(* IEC 61131-3 sources: Test-Git_ESME26/TestProgettoESME_26.fbsproj/AxisModuleLib Migration/DiagSource, 7 files *)

(* ---- AXM_FC_EtCamTypeToString.fn.st ---- *)
FUNCTION INTERNAL AXM_FC_EtCamTypeToString : STRING[80]
VAR_INPUT
	i_etCamType	: CMT.ET_CamType;
END_VAR
VAR
END_VAR

CASE i_etCamType OF
	CMT.ET_CamType.Straight:
		AXM_FC_EtCamTypeToString := 'Straight';

	CMT.ET_CamType.Poly5Com:
		AXM_FC_EtCamTypeToString := 'Poly5Com';

	CMT.ET_CamType.SimplSin:
		AXM_FC_EtCamTypeToString := 'SimplSin';

	CMT.ET_CamType.IncliSin:
		AXM_FC_EtCamTypeToString := 'IncliSin';

	CMT.ET_CamType.ModiSin:
		AXM_FC_EtCamTypeToString := 'ModiSin';

	CMT.ET_CamType.ModAccTr:
		AXM_FC_EtCamTypeToString := 'ModAccTr';

	CMT.ET_CamType.Poly5:
		AXM_FC_EtCamTypeToString := 'Poly5';

	CMT.ET_CamType.Parable2:
		AXM_FC_EtCamTypeToString := 'Parable2';

	CMT.ET_CamType.UserCam:
		AXM_FC_EtCamTypeToString := 'UserCam';

	CMT.ET_CamType.ModiSinCom:
		AXM_FC_EtCamTypeToString := 'ModiSinCom';

	CMT.ET_CamType.ModAccTrCom:
		AXM_FC_EtCamTypeToString := 'ModAccTrCom';

	CMT.ET_CamType.HarmoComb:
		AXM_FC_EtCamTypeToString := 'HarmoComb';

	CMT.ET_CamType.SinStraightComb:
		AXM_FC_EtCamTypeToString := 'SinStraightComb';

ELSE
	AXM_FC_EtCamTypeToString := Standard.CONCAT('Unknown CamType ', INT_TO_STRING(i_etCamType));
END_CASE

(* ---- AXM_FC_EtHomeModeToString.fn.st ---- *)
FUNCTION INTERNAL AXM_FC_EtHomeModeToString : STRING[80]
VAR_INPUT
	i_etHomeMode : PDL_ET_HomeMode;
END_VAR
VAR
END_VAR

AXM_FC_EtHomeModeToString := TO_STRING(i_etHomeMode);

(* ---- AXM_FC_EtMultiCamCsModeMasterToString.fn.st ---- *)
FUNCTION AXM_FC_EtMultiCamCsModeMasterToString : STRING[80]
VAR_INPUT
	i_etCsModeMaster	: PDL_ET_MultiCamCsModeMaster;
END_VAR
VAR
END_VAR

AXM_FC_EtMultiCamCsModeMasterToString := TO_STRING(i_etCsModeMaster);

(* ---- AXM_FC_EtMultiCamCsModeSlaveToString.fn.st ---- *)
FUNCTION AXM_FC_EtMultiCamCsModeSlaveToString : STRING[80]
VAR_INPUT
	i_etCsModeSlave	: PDL_ET_MultiCamCsModeSlave;
END_VAR
VAR
END_VAR

AXM_FC_EtMultiCamCsModeSlaveToString := To_string(i_etCsModeSlave);

(* ---- AXM_FC_EtMultiCamWsModeToString.fn.st ---- *)
FUNCTION AXM_FC_EtMultiCamWsModeToString : STRING[80]
VAR_INPUT
	i_etWsMode	: PDL_ET_MultiCamWsMode;
END_VAR
VAR
END_VAR

CASE i_etWsMode OF
	PDL_ET_MultiCamWsMode.StoredCamMoveAlwaysNoPositionCheck:
		AXM_FC_EtMultiCamWsModeToString := 'StoredCamMoveAlwaysNoPositionCheck';

	PDL_ET_MultiCamWsMode.StoredCamMoveToCamPositonInWsWindow:
		AXM_FC_EtMultiCamWsModeToString := 'StoredCamMoveToCamPositonInWsWindow';

	PDL_ET_MultiCamWsMode.StoredCamMoveForwardToCamPositon:
		AXM_FC_EtMultiCamWsModeToString := 'StoredCamMoveForwardToCamPositon';

	PDL_ET_MultiCamWsMode.StoredCamMoveBackwardToCamPosition:
		AXM_FC_EtMultiCamWsModeToString := 'StoredCamMoveBackwardToCamPosition';

	PDL_ET_MultiCamWsMode.StoredCamShowCamPosition:
		AXM_FC_EtMultiCamWsModeToString := 'StoredCamShowCamPosition';

	PDL_ET_MultiCamWsMode.StoredCamSetMasterPositionToRelatedSlavePosition:
		AXM_FC_EtMultiCamWsModeToString := 'StoredCamSetMasterPositionToRelatedSlavePosition';

	PDL_ET_MultiCamWsMode.NewCamMoveAlwaysNoPositionCheck:
		AXM_FC_EtMultiCamWsModeToString := 'NewCamMoveAlwaysNoPositionCheck';

	PDL_ET_MultiCamWsMode.NewCamMoveToCamPositonInWsWindow:
		AXM_FC_EtMultiCamWsModeToString := 'NewCamMoveToCamPositonInWsWindow';

	PDL_ET_MultiCamWsMode.NewCamMoveForwardToCamPositon:
		AXM_FC_EtMultiCamWsModeToString := 'NewCamMoveForwardToCamPositon';

	PDL_ET_MultiCamWsMode.NewCamMoveBackwardToCamPosition:
		AXM_FC_EtMultiCamWsModeToString := 'NewCamMoveBackwardToCamPosition';

	PDL_ET_MultiCamWsMode.NewCamShowCamPosition:
		AXM_FC_EtMultiCamWsModeToString := 'NewCamShowCamPosition';

	PDL_ET_MultiCamWsMode.NewCamSetMasterPositionToRelatedSlavePosition:
		AXM_FC_EtMultiCamWsModeToString := 'NewCamSetMasterPositionToRelatedSlavePosition';

	ELSE
		AXM_FC_EtMultiCamWsModeToString := Standard.CONCAT('Unknown WsMode ', INT_TO_STRING(i_etWsMode));
END_CASE

(* ---- AXM_FC_EtPosModeToString.fn.st ---- *)
FUNCTION AXM_FC_EtPosModeToString : STRING[80]
VAR_INPUT
	i_etPosMode	: PDL_ET_PosMode;
END_VAR
VAR
END_VAR

AXM_FC_EtPosModeToString := TO_STRING(i_etPosMode);

(* ---- AXM_FB_AxisModuleDiagSource.fb.st ---- *)
FUNCTION_BLOCK PUBLIC AXM_FB_AxisModuleDiagSource
VAR_INPUT
	i_xEnable			: BOOL;
	i_xDiagQuit			: BOOL;
	i_xPrintCamData		: BOOL := TRUE;
END_VAR
VAR_IN_OUT
	iq_stComStructure	: TPL.ST_DiagnosticsManagerToDiagSource;
	iq_stMachineItf		: TPL.ST_StandardModuleInterface;
END_VAR
VAR_OUTPUT
	q_xActive			: BOOL;
	q_xReady			: BOOL;
	q_etDiag			: GD.ET_Diag := GD.ET_Diag.Ok;
	q_etDiagExt			: AXM_ET_DiagExt := AXM_ET_DiagExt.Disabled;
	q_sMsg				: STRING[80];
END_VAR
VAR
	xEnableFlag		: BOOL;
	diState			: DINT;
	udiOwnSourceId	: UDINT := 0;
	fbTreeWriter	: TPL.FB_TreeWriter;
	diOldCmd		: DINT := 0;
	diCmdExecState	: DINT := 0;
	lrSumNodes		: LREAL := 1;
	pstTmp			: POINTER TO TPL.ST_StandardModuleInterface;
	audiHierarchy	: ARRAY[1..c_udiMaxLevel] OF UDINT;
	udiLevelCounter	: UDINT := 1;
	apstHierarchy	: ARRAY[1..c_udiMaxLevel] OF POINTER TO TPL.ST_StandardModuleInterface;
	xLoop			: BOOL;
	pstInterface	: POINTER TO AXM_ST_ModuleInterface;
	pdw				: POINTER TO TPL.TYPE_ADDRESS;
	sTmp			: STRING[80];
	diMotionParCounter	: DINT;
	diCamPointCounter	: DINT;
	diCount			: DINT;
	pstChar			: POINTER TO STRING;
	sModuleMain		: STRING[80];
	sModuleName		: STRING;
	diLoopBreaker	: DINT;
	etDiag			: GD.ET_Diag;
	etDiagExtTPL	: TPL.ET_DiagExt;
	sMsg			: STRING[80];
	rtrigDiagQuit	: Standard.R_TRIG;
END_VAR
VAR CONSTANT
	c_sName			: STRING[TPL.Gc_udiTableWriterMaxNameLength] := 'AxisModule_Interface' ;
	c_sTypeName		: STRING[TPL.Gc_udiTableWriterMaxNameLength] := 'AXM_Interface' ;
	c_udiMaxLevel	: UDINT := 8;
END_VAR

IF i_xEnable AND NOT xEnableFlag THEN
	xEnableFlag := TRUE;

	q_xActive := TRUE;

	SetDiagOutputs(	i_etDiag	:= GD.ET_Diag.Ok,
					i_etDiagExt	:= AXM_ET_DiagExt.WaitUntilDiagnosticsManagerReady,
					i_sMsg		:= '');
	diState := 10;

ELSIF NOT i_xEnable AND xEnableFlag THEN
	xEnableFlag := FALSE;

	IF udiOwnSourceId <> 0 THEN
		SetDiagOutputs(	i_etDiag	:= GD.ET_Diag.Ok,
						i_etDiagExt	:= AXM_ET_DiagExt.WaitUntilDisabled,
						i_sMsg		:= '');
		diState := 100;

	ELSIF udiOwnSourceId = 0 THEN
		SetDiagOutputs(	i_etDiag	:= GD.ET_Diag.Ok,
						i_etDiagExt	:= AXM_ET_DiagExt.Disabled,
						i_sMsg		:= '');
	END_IF
END_IF

DiagQuit();

CASE diState OF

	0:	(* Disable & exception state *)

	10:	(* Wait until diagnostics manager ready *)
		IF iq_stComStructure.i_xDiagnosticsManagerReady THEN

			SetDiagOutputs(	i_etDiag	:= GD.ET_Diag.Ok,
							i_etDiagExt	:= AXM_ET_DiagExt.WaitUntilDiagSourceRegistered,
							i_sMsg		:= '');
			diState := 20;
		END_IF

	20:	(* Wait until diag source registered *)
		IF NOT iq_stComStructure.i_xDiagnosticsManagerReady THEN

			SetDiagOutputs(	i_etDiag	:= GD.ET_Diag.Ok,
							i_etDiagExt	:= AXM_ET_DiagExt.WaitUntilDiagnosticsManagerReady,
							i_sMsg		:= '');
			diState := 10;
			RETURN;

		(* only write to register structure if no one else has done it in this cylce *)
		ELSIF (NOT iq_stComStructure.iq_stRegister.xUsed AND iq_stComStructure.iq_stRegister.udiNextId <> 0) THEN
			(* register *)
			iq_stComStructure.iq_stRegister.xUsed := TRUE;

			iq_stComStructure.iq_stRegister.sName		:= c_sName;
			iq_stComStructure.iq_stRegister.sTypeName	:= c_sTypeName;

			udiOwnSourceId := iq_stComStructure.iq_stRegister.udiNextId; (* register with this id; required for the following communication *)
		ELSE
			RETURN;
		END_IF

		q_xReady := TRUE;

		SetDiagOutputs(	i_etDiag	:= GD.ET_Diag.Ok,
						i_etDiagExt	:= AXM_ET_DiagExt.WaitForCommunication,
						i_sMsg		:= '');
		diState := 30;

	30:	(* Wait for communication *)
		IF NOT iq_stComStructure.i_xDiagnosticsManagerReady THEN

			CancelWriting();

			udiOwnSourceId	:= 0;

			SetDiagOutputs(	i_etDiag	:= GD.ET_Diag.Ok,
							i_etDiagExt	:= AXM_ET_DiagExt.WaitUntilDiagnosticsManagerReady,
							i_sMsg		:= '');
			diState := 10;
			RETURN;

		ELSIF (iq_stComStructure.i_udiComWithId = udiOwnSourceId) THEN		(* Am I adressed? *)

			WriteDiagDataControl();

		ELSE
			iq_stComStructure.q_lrProgress := 0.0;

			CancelWriting();

			SetDiagOutputs(	i_etDiag	:= GD.ET_Diag.Ok,
							i_etDiagExt	:= AXM_ET_DiagExt.WaitForCommunication,
							i_sMsg		:= '');
		END_IF

	100: (* Wait until disabled *)
		IF NOT iq_stComStructure.i_xDiagnosticsManagerReady THEN

			CancelWriting();

			udiOwnSourceId	:= 0;

			SetDiagOutputs(	i_etDiag	:= GD.ET_Diag.Ok,
							i_etDiagExt	:= AXM_ET_DiagExt.Disabled,
							i_sMsg		:= '');

		ELSIF (iq_stComStructure.i_udiComWithId = udiOwnSourceId) THEN		(* Am I adressed? *)

			WriteDiagDataControl();

		(* only write to register structure if no one else has done it in this cylce *)
		ELSIF (NOT iq_stComStructure.iq_stRegister.xUsed AND NOT iq_stComStructure.iq_stRegister.xUnsubscribe) AND
			   NOT iq_stComStructure.i_xDiagnosticsActive THEN

			iq_stComStructure.iq_stRegister.xUsed			:= TRUE;

			iq_stComStructure.iq_stRegister.xUnsubscribe	:= TRUE;
			iq_stComStructure.iq_stRegister.udiSourceId		:= udiOwnSourceId;

			q_xActive := FALSE;

			SetDiagOutputs(	i_etDiag	:= GD.ET_Diag.Ok,
							i_etDiagExt	:= AXM_ET_DiagExt.Disabled,
							i_sMsg		:= '');
		END_IF
END_CASE

IF q_xActive THEN
	IF(diCmdExecState <> 0) THEN
		WriteDiagDataToFile();

		IF(iq_stComStructure.iq_diCmd <= 0) THEN
			diOldCmd := iq_stComStructure.iq_diCmd;
		END_IF
	END_IF
END_IF
